FUNCTION_BLOCK TankResis (* Composite Function Block Type *)
  (* Standard: 61499-2 *)
  (* Version 0.0, 6/21/2016, Andrei, nxtControl GmbH, template *)
  PACKAGE Main;
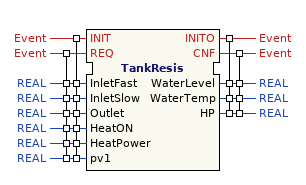
  EVENT_INPUT
    INIT WITH InletFast, InletSlow, Outlet, HeatON, HeatPower, pv1; (* Initialization Request *)
    REQ WITH InletFast, InletSlow, Outlet, HeatON, HeatPower, pv1; (* Normal Execution Request *)
  END_EVENT
  EVENT_OUTPUT
    INITO WITH WaterLevel, WaterTemp, HP; (* Initialization Confirm *)
    CNF WITH WaterLevel, WaterTemp, HP; (* Execution Confirmation *)
  END_EVENT
  VAR_INPUT
    InletFast : REAL; (* Input event qualifier *)
    InletSlow : REAL;
    Outlet : REAL;
    HeatON : REAL;
    HeatPower : REAL;
    pv1 : REAL;
  END_VAR
  VAR_OUTPUT
    WaterLevel : REAL; (* Output event qualifier *)
    WaterTemp : REAL;
    HP : REAL;
  END_VAR
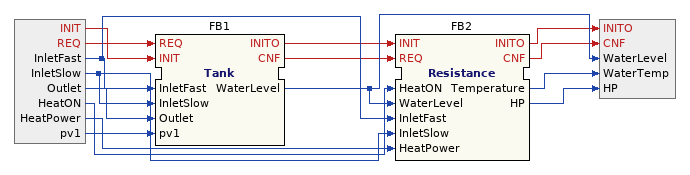
  FBS
    FB1 : Tank;
    FB2 : Resistance;
  END_FBS
  EVENT_CONNECTIONS
    REQ TO FB1.REQ;
    INIT TO FB1.INIT;
    FB1.INITO TO FB2.INIT;
    FB1.CNF TO FB2.REQ;
    FB2.INITO TO INITO;
    FB2.CNF TO CNF;
  END_CONNECTIONS
  DATA_CONNECTIONS
    InletFast TO FB1.InletFast;
    InletSlow TO FB1.InletSlow;
    Outlet TO FB1.Outlet;
    HeatON TO FB2.HeatON;
    FB1.WaterLevel TO FB2.WaterLevel;
    FB2.Temperature TO WaterTemp;
    FB1.WaterLevel TO WaterLevel;
    InletFast TO FB2.InletFast;
    InletSlow TO FB2.InletSlow;
    HeatPower TO FB2.HeatPower;
    pv1 TO FB1.pv1;
    FB2.HP TO HP;
  END_CONNECTIONS
END_FUNCTION_BLOCK
